(* IEC 61131-3 sources: llm-plc-st-eval/data/processed_definitivo/claude-sonnet-4-6/I1/zero_shot, 3 files *)

(* ---- ejec_1.st ---- *)
FUNCTION_BLOCK FB_Semaforo
VAR_INPUT
    habilitado : BOOL; (* Habilita la secuencia normal del semáforo *)
END_VAR

VAR_OUTPUT
    luzV : BOOL; (* Luz verde *)
    luzA : BOOL; (* Luz amarilla *)
    luzR : BOOL; (* Luz roja *)
END_VAR

VAR
    (* Temporizadores TON estándar IEC 61131-3 *)
    tVerde      : TON; (* Temporizador fase verde:   20 s *)
    tAmarillo   : TON; (* Temporizador fase amarilla: 4 s *)
    tRojo       : TON; (* Temporizador fase roja:    15 s *)
    tParpadeo   : TON; (* Temporizador parpadeo:      1 s *)

    (* Estado de la máquina de estados *)
    (* 0 = Verde, 1 = Amarillo, 2 = Rojo, 3 = Amarillo intermitente *)
    estado      : INT := 0;

    (* Bit auxiliar para el parpadeo del amarillo intermitente *)
    parpadeoOn  : BOOL := FALSE;
END_VAR

(* ─────────────────────────────────────────────────────────────────────────── *)
(*  Lógica principal                                                           *)
(* ─────────────────────────────────────────────────────────────────────────── *)

IF NOT habilitado THEN
    (* ── Modo amarillo intermitente ─────────────────────────────────────── *)

    (* Si veníamos de la secuencia normal, reiniciamos al estado intermitente *)
    IF estado <> 3 THEN
        estado     := 3;
        parpadeoOn := FALSE;
        (* Apagar temporizadores de secuencia normal *)
        tVerde(IN := FALSE, PT := T#20S);
        tAmarillo(IN := FALSE, PT := T#4S);
        tRojo(IN := FALSE, PT := T#15S);
        (* Arrancar temporizador de parpadeo *)
        tParpadeo(IN := FALSE, PT := T#1S);
    END_IF;

    (* Temporizador de parpadeo: alterna cada 1 s *)
    tParpadeo(IN := TRUE, PT := T#1S);
    IF tParpadeo.Q THEN
        parpadeoOn := NOT parpadeoOn; (* Invertir estado del parpadeo *)
        tParpadeo(IN := FALSE, PT := T#1S); (* Reiniciar temporizador *)
    END_IF;

    (* Salidas: solo amarillo parpadea, verde y rojo apagados *)
    luzV := FALSE;
    luzA := parpadeoOn;
    luzR := FALSE;

ELSE
    (* ── Secuencia normal cíclica ────────────────────────────────────────── *)

    (* Si veníamos del modo intermitente, reiniciar en verde *)
    IF estado = 3 THEN
        estado := 0;
        parpadeoOn := FALSE;
        tParpadeo(IN := FALSE, PT := T#1S); (* Detener parpadeo *)
    END_IF;

    CASE estado OF

        0: (* ── VERDE 20 s ─────────────────────────────────────────────── *)
            tVerde(IN := TRUE, PT := T#20S);
            luzV := TRUE;
            luzA := FALSE;
            luzR := FALSE;
            IF tVerde.Q THEN
                tVerde(IN := FALSE, PT := T#20S); (* Reiniciar temporizador *)
                estado := 1;                       (* Pasar a amarillo *)
            END_IF;

        1: (* ── AMARILLO 4 s ────────────────────────────────────────────── *)
            tAmarillo(IN := TRUE, PT := T#4S);
            luzV := FALSE;
            luzA := TRUE;
            luzR := FALSE;
            IF tAmarillo.Q THEN
                tAmarillo(IN := FALSE, PT := T#4S); (* Reiniciar temporizador *)
                estado := 2;                         (* Pasar a rojo *)
            END_IF;

        2: (* ── ROJO 15 s ───────────────────────────────────────────────── *)
            tRojo(IN := TRUE, PT := T#15S);
            luzV := FALSE;
            luzA := FALSE;
            luzR := TRUE;
            IF tRojo.Q THEN
                tRojo(IN := FALSE, PT := T#15S); (* Reiniciar temporizador *)
                estado := 0;                      (* Volver a verde *)
            END_IF;

        ELSE
            (* Estado inesperado: forzar reinicio en verde *)
            estado := 0;

    END_CASE;

END_IF;

(* ---- ejec_2.st ---- *)
FUNCTION_BLOCK FB_Semaforo
VAR_INPUT
    habilitado : BOOL; (* Habilita la secuencia normal del semáforo *)
END_VAR

VAR_OUTPUT
    luzV : BOOL; (* Luz verde *)
    luzA : BOOL; (* Luz amarilla *)
    luzR : BOOL; (* Luz roja *)
END_VAR

VAR
    (* Temporizadores para cada fase de la secuencia normal *)
    tVerde    : TON; (* Temporiza la fase verde  - 20 s *)
    tAmarillo : TON; (* Temporiza la fase amarilla - 4 s *)
    tRojo     : TON; (* Temporiza la fase roja   - 15 s *)

    (* Temporizador para el amarillo intermitente *)
    tIntermitente : TON; (* Temporiza cada semiciclo de 1 s *)

    (* Estado interno de la secuencia normal *)
    (* 0 = Verde, 1 = Amarillo, 2 = Rojo *)
    estado : INT := 0;

    (* Bit de parpadeo para el amarillo intermitente *)
    parpadeo : BOOL := FALSE;
END_VAR

(* ─────────────────────────────────────────────────────────────
   Lógica principal
   ───────────────────────────────────────────────────────────── *)

IF NOT habilitado THEN
    (* ── Modo amarillo intermitente ─────────────────────────── *)

    (* Reiniciar temporizadores de secuencia normal *)
    tVerde(IN    := FALSE, PT := T#20S);
    tAmarillo(IN := FALSE, PT := T#4S);
    tRojo(IN     := FALSE, PT := T#15S);

    (* Reiniciar estado para que al habilitar arranque en verde *)
    estado := 0;

    (* Temporizador de 1 s para el parpadeo *)
    tIntermitente(IN := TRUE, PT := T#1S);

    IF tIntermitente.Q THEN
        (* Conmutar el bit de parpadeo y reiniciar el temporizador *)
        parpadeo          := NOT parpadeo;
        tIntermitente(IN  := FALSE, PT := T#1S); (* Reset *)
        tIntermitente(IN  := TRUE,  PT := T#1S); (* Rearranque *)
    END_IF;

    (* Salidas: solo amarillo parpadea *)
    luzV := FALSE;
    luzA := parpadeo;
    luzR := FALSE;

ELSE
    (* ── Modo secuencia normal ───────────────────────────────── *)

    (* Detener y resetear el temporizador de intermitente *)
    tIntermitente(IN := FALSE, PT := T#1S);
    parpadeo := FALSE;

    CASE estado OF

        0: (* ── Verde ── *)
            luzV := TRUE;
            luzA := FALSE;
            luzR := FALSE;

            tVerde(IN := TRUE, PT := T#20S);

            IF tVerde.Q THEN
                tVerde(IN := FALSE, PT := T#20S); (* Reset *)
                estado := 1;                       (* Pasar a amarillo *)
            END_IF;

        1: (* ── Amarillo ── *)
            luzV := FALSE;
            luzA := TRUE;
            luzR := FALSE;

            tAmarillo(IN := TRUE, PT := T#4S);

            IF tAmarillo.Q THEN
                tAmarillo(IN := FALSE, PT := T#4S); (* Reset *)
                estado := 2;                         (* Pasar a rojo *)
            END_IF;

        2: (* ── Rojo ── *)
            luzV := FALSE;
            luzA := FALSE;
            luzR := TRUE;

            tRojo(IN := TRUE, PT := T#15S);

            IF tRojo.Q THEN
                tRojo(IN := FALSE, PT := T#15S); (* Reset *)
                estado := 0;                      (* Volver a verde *)
            END_IF;

        ELSE
            (* Estado inválido: reiniciar en verde *)
            estado := 0;

    END_CASE;

END_IF;

(* ---- ejec_3.st ---- *)
FUNCTION_BLOCK FB_Semaforo
VAR_INPUT
    habilitado : BOOL; (* Habilita la secuencia normal del semáforo *)
END_VAR

VAR_OUTPUT
    luzV : BOOL; (* Luz verde *)
    luzA : BOOL; (* Luz amarilla *)
    luzR : BOOL; (* Luz roja *)
END_VAR

VAR
    (* Temporizadores para cada fase *)
    tVerde     : TON; (* Temporizador fase verde  - 20 s *)
    tAmarillo  : TON; (* Temporizador fase amarilla - 4 s *)
    tRojo      : TON; (* Temporizador fase roja   - 15 s *)
    tBlink     : TON; (* Temporizador parpadeo amarillo - 1 s *)

    (* Estado de la secuencia normal *)
    (* 0 = Verde, 1 = Amarillo, 2 = Rojo *)
    estado     : INT := 0;

    (* Estado interno del parpadeo (TRUE = encendido, FALSE = apagado) *)
    blinkOn    : BOOL := FALSE;
END_VAR

(* ─────────────────────────────────────────────────────────────────────────── *)

IF NOT habilitado THEN
    (* ── Modo amarillo intermitente ─────────────────────────────────────── *)

    (* Reiniciar temporizadores de secuencia normal *)
    tVerde(IN := FALSE);
    tAmarillo(IN := FALSE);
    tRojo(IN := FALSE);

    (* Reiniciar estado para que al habilitar arranque en verde *)
    estado := 0;

    (* Temporizador de parpadeo: ciclo de 1 s *)
    tBlink(IN := TRUE, PT := T#1S);

    IF tBlink.Q THEN
        (* Conmutar estado del parpadeo y reiniciar temporizador *)
        blinkOn := NOT blinkOn;
        tBlink(IN := FALSE); (* Reset del temporizador *)
    END_IF;

    (* Asignar salidas: solo amarillo parpadea *)
    luzV := FALSE;
    luzA := blinkOn;
    luzR := FALSE;

ELSE
    (* ── Modo secuencia normal ───────────────────────────────────────────── *)

    (* Detener y resetear temporizador de parpadeo *)
    tBlink(IN := FALSE);
    blinkOn := FALSE;

    CASE estado OF

        0: (* ── Fase VERDE ── *)
            luzV := TRUE;
            luzA := FALSE;
            luzR := FALSE;

            tVerde(IN := TRUE, PT := T#20S);

            IF tVerde.Q THEN
                tVerde(IN := FALSE); (* Reset temporizador *)
                estado := 1;         (* Pasar a amarillo *)
            END_IF;

        1: (* ── Fase AMARILLA ── *)
            luzV := FALSE;
            luzA := TRUE;
            luzR := FALSE;

            tAmarillo(IN := TRUE, PT := T#4S);

            IF tAmarillo.Q THEN
                tAmarillo(IN := FALSE); (* Reset temporizador *)
                estado := 2;            (* Pasar a rojo *)
            END_IF;

        2: (* ── Fase ROJA ── *)
            luzV := FALSE;
            luzA := FALSE;
            luzR := TRUE;

            tRojo(IN := TRUE, PT := T#15S);

            IF tRojo.Q THEN
                tRojo(IN := FALSE); (* Reset temporizador *)
                estado := 0;        (* Volver a verde *)
            END_IF;

        ELSE
            (* Estado inválido: reiniciar en verde *)
            estado := 0;

    END_CASE;

END_IF;
